Fanuc KAREL source: ks00038.KL

PROGRAM KS00038
%STACKSIZE=65535
%PRIORITY=65535
%NOLOCKGROUP
VAR
A : ARRAY[4] OF POSITION
B : ARRAY[4] OF POSITION
FLAG : BOOLEAN
N : INTEGER
STATUS : INTEGER
PN : STRING[80]
VN : STRING[80]
BEGIN
PN=''
VN='A'
-- UNRESOLVED_PC line 19 opcodes [22 22 1E] marker_code=27
END KS00038
